Fanuc KAREL source: NC0001.compact.KL

PROGRAM NC0001
%STACKSIZE=65535
%PRIORITY=65535
%NOLOCKGROUP
ROUTINE R FROM NC0001
ROUTINE R
VAR
S1 : INTEGER
BEGIN
S1=1
S1=(S1 + 1)
END R
BEGIN
R
END NC0001
